{attribute 'Tc2GvlVarNames'}
VAR_GLOBAL
	stgGr00Alarm			:ST_AlarmRef;
END_VAR

(* stored: Version 1.1.0.1, ProductVersion 3.1.4024.15
   GVL GVL_Gr00Alarm: Id {76050387-16fd-412f-9370-dcd4cacdfa63} *)
